{attribute 'qualified_only'}
{attribute 'strict'}
TYPE HmiCommandCode :
(
	NONE := 0,
	MANUAL_DRIVE,
	START_MAPPING,
	START_SWEEPING,
	PAUSE,
	RESUME,
	STOP,
	GO_TO_DOCK,
	EMERGENCY_STOP,
	RESET,
	SET_POSE
) INT;
END_TYPE

(* stored: Version 1.1.0.1, ProductVersion 3.1.4026.12
   DUT HmiCommandCode: Id {0f7c0614-0470-5b09-aa78-6db22868f2a3} *)
